FUNCTION_BLOCK Subestacao (* Subestacao / QGBT e geradores - ETE Tijuco Preto *)
  (* Standard: 61499-2 *)
  (* Version 1.2, 11/11/2026, Hidryco, Hidryco, 1.2: disjuntores ligados do PCE LODO (900) lidos pelo M262_Substacao na remota 1 do Lodo (.135): ${PATH}dj900_* e ${PATH}stsFalhaRemotaLODO -> IThis DJ_900_* e FALHA_REMOTA_LODO (PCE com logica invertida). 1.0: QGBT 440 V da ETE Tijuco Preto (unifilar HID-PE-DE-ETE-ELE-002): QTAM 1 (G2) -> 1Q1 -> barra A, QTAM 2 (G1) -> 1Q2 -> barra B, 1Q0 acoplamento. Disjuntores pelos DIs da remota 1 (A3/A4/A5 TM3DI32K do PCE SUBESTACAO) publicados por IO_DI32 em ${PATH}dj<nome>, ${PATH}mp<sinal>_1q<n> e ${PATH}stsFalhaRemota1. Geradores pelos Gerador_Generico internos GMG_G1 (QTAM 2) e GMG_G2 (QTAM 1). Cargas liberadas no gerador escolhidas na IHM (persistentes, padrao liberado): saidas HAB_* e stsPlantaNoGerador para os CATs de processo. v1.1: comandos de abrir/fechar dos Masterpact pela IHM (fpComandos) com intertravamentos, publicados em ${PATH}cmdAbrir1q1 ... ${PATH}cmdFechar1q2 para o IO_DQ32 do A8 TM3DQ32TK da remota 1 (word 0 b05..b10, escrita pelo M262_Substacao); reservas no unifilar. *)
  PACKAGE Hidryco.HidrycoLib;
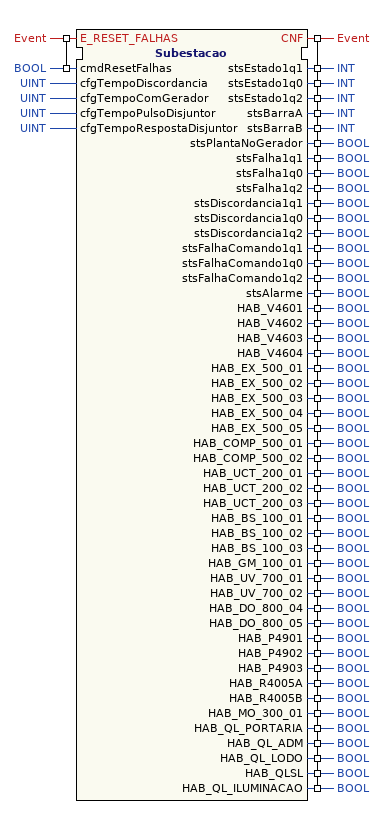
  EVENT_INPUT
    E_RESET_FALHAS WITH cmdResetFalhas; (* Reconhecimento pelo processo com cmdResetFalhas = TRUE *)
  END_EVENT
  EVENT_OUTPUT
    CNF WITH stsEstado1q1, stsEstado1q0, stsEstado1q2, stsBarraA, stsBarraB, stsPlantaNoGerador, stsFalha1q1, stsFalha1q0, stsFalha1q2, stsDiscordancia1q1, stsDiscordancia1q0, stsDiscordancia1q2, stsFalhaComando1q1, stsFalhaComando1q0, stsFalhaComando1q2, stsAlarme, HAB_V4601, HAB_V4602, HAB_V4603, HAB_V4604, HAB_EX_500_01, HAB_EX_500_02, HAB_EX_500_03, HAB_EX_500_04, HAB_EX_500_05, HAB_COMP_500_01, HAB_COMP_500_02, HAB_UCT_200_01, HAB_UCT_200_02, HAB_UCT_200_03, HAB_BS_100_01, HAB_BS_100_02, HAB_BS_100_03, HAB_GM_100_01, HAB_UV_700_01, HAB_UV_700_02, HAB_DO_800_04, HAB_DO_800_05, HAB_P4901, HAB_P4902, HAB_P4903, HAB_R4005A, HAB_R4005B, HAB_MO_300_01, HAB_QL_PORTARIA, HAB_QL_ADM, HAB_QL_LODO, HAB_QLSL, HAB_QL_ILUMINACAO; (* Estados do QGBT e cargas liberadas no gerador (so na mudanca) *)
  END_EVENT
  VAR_INPUT
    cmdResetFalhas : BOOL; (* TRUE = reconhecimento (com o evento E_RESET_FALHAS) *)
    cfgTempoDiscordancia : UINT := 5; (* Tempo (s) com aberto/fechado discordantes para o aviso de posicao indefinida *)
    cfgTempoComGerador : UINT := 10; (* Tempo (s) sem comunicacao com os AGC 150 para confirmar a falha *)
    cfgTempoPulsoDisjuntor : UINT := 1; (* Tempo (s) do pulso de abrir/fechar dos Masterpact (o pulso acaba antes se o disjuntor mudar de estado) *)
    cfgTempoRespostaDisjuntor : UINT := 5; (* Tempo (s) para o Masterpact mudar de estado depois do comando (senao: aviso de sem resposta) *)
  END_VAR
  VAR_OUTPUT
    stsEstado1q1 : INT; (* Disjuntor 1Q1: 0 indefinido (sem comunicacao), 1 aberto, 2 fechado, 3 discordante *)
    stsEstado1q0 : INT; (* Disjuntor 1Q0: 0 indefinido (sem comunicacao), 1 aberto, 2 fechado, 3 discordante *)
    stsEstado1q2 : INT; (* Disjuntor 1Q2: 0 indefinido (sem comunicacao), 1 aberto, 2 fechado, 3 discordante *)
    stsBarraA : INT; (* Fonte da barra A (1Q1): 0 sem alimentacao, 1 rede, 2 gerador, 3 indefinida *)
    stsBarraB : INT; (* Fonte da barra B (1Q2): 0 sem alimentacao, 1 rede, 2 gerador, 3 indefinida *)
    stsPlantaNoGerador : BOOL; (* Alguma QTAM com o disjuntor do gerador fechado (planta nos geradores) *)
    stsFalha1q1 : BOOL; (* Disjuntor 1Q1 em falha (desarmado) *)
    stsFalha1q0 : BOOL; (* Disjuntor 1Q0 em falha (desarmado) *)
    stsFalha1q2 : BOOL; (* Disjuntor 1Q2 em falha (desarmado) *)
    stsDiscordancia1q1 : BOOL; (* Disjuntor 1Q1: posição indefinida (aberto e fechado discordantes) *)
    stsDiscordancia1q0 : BOOL; (* Disjuntor 1Q0: posição indefinida (aberto e fechado discordantes) *)
    stsDiscordancia1q2 : BOOL; (* Disjuntor 1Q2: posição indefinida (aberto e fechado discordantes) *)
    stsFalhaComando1q1 : BOOL; (* Disjuntor 1Q1 não respondeu ao comando de abrir/fechar *)
    stsFalhaComando1q0 : BOOL; (* Disjuntor 1Q0 não respondeu ao comando de abrir/fechar *)
    stsFalhaComando1q2 : BOOL; (* Disjuntor 1Q2 não respondeu ao comando de abrir/fechar *)
    stsAlarme : BOOL; (* Algum alarme do QGBT *)
    HAB_V4601 : BOOL; (* V4601 - Soprador 01 liberado para operar com a planta nos geradores *)
    HAB_V4602 : BOOL; (* V4602 - Soprador 02 liberado para operar com a planta nos geradores *)
    HAB_V4603 : BOOL; (* V4603 - Soprador 03 liberado para operar com a planta nos geradores *)
    HAB_V4604 : BOOL; (* V4604 - Soprador 04 liberado para operar com a planta nos geradores *)
    HAB_EX_500_01 : BOOL; (* 500-EX-01 - Exaustor 01 liberado para operar com a planta nos geradores *)
    HAB_EX_500_02 : BOOL; (* 500-EX-02 - Exaustor 02 liberado para operar com a planta nos geradores *)
    HAB_EX_500_03 : BOOL; (* 500-EX-03 - Exaustor 03 liberado para operar com a planta nos geradores *)
    HAB_EX_500_04 : BOOL; (* 500-EX-04 - Exaustor 04 liberado para operar com a planta nos geradores *)
    HAB_EX_500_05 : BOOL; (* 500-EX-05 - Exaustor 05 liberado para operar com a planta nos geradores *)
    HAB_COMP_500_01 : BOOL; (* 500-COMP-01 - Compressor 01 liberado para operar com a planta nos geradores *)
    HAB_COMP_500_02 : BOOL; (* 500-COMP-02 - Compressor 02 liberado para operar com a planta nos geradores *)
    HAB_UCT_200_01 : BOOL; (* 200-UCT-01 - Unid. compacta 01 liberado para operar com a planta nos geradores *)
    HAB_UCT_200_02 : BOOL; (* 200-UCT-02 - Unid. compacta 02 liberado para operar com a planta nos geradores *)
    HAB_UCT_200_03 : BOOL; (* 200-UCT-03 - Unid. compacta 03 liberado para operar com a planta nos geradores *)
    HAB_BS_100_01 : BOOL; (* 100-BS-01 - Bomba 01 liberado para operar com a planta nos geradores *)
    HAB_BS_100_02 : BOOL; (* 100-BS-02 - Bomba 02 liberado para operar com a planta nos geradores *)
    HAB_BS_100_03 : BOOL; (* 100-BS-03 - Bomba 03 liberado para operar com a planta nos geradores *)
    HAB_GM_100_01 : BOOL; (* 100-GM-01 - Grade mecanizada liberado para operar com a planta nos geradores *)
    HAB_UV_700_01 : BOOL; (* 700-UV-01 - Sistema UV 01 liberado para operar com a planta nos geradores *)
    HAB_UV_700_02 : BOOL; (* 700-UV-02 - Sistema UV 02 liberado para operar com a planta nos geradores *)
    HAB_DO_800_04 : BOOL; (* 800-DO-04 - Bomba dosadora 04 liberado para operar com a planta nos geradores *)
    HAB_DO_800_05 : BOOL; (* 800-DO-05 - Bomba dosadora 05 liberado para operar com a planta nos geradores *)
    HAB_P4901 : BOOL; (* P4901 - Bomba submersível 01 liberado para operar com a planta nos geradores *)
    HAB_P4902 : BOOL; (* P4902 - Bomba submersível 02 liberado para operar com a planta nos geradores *)
    HAB_P4903 : BOOL; (* P4903 - Bomba submersível 03 liberado para operar com a planta nos geradores *)
    HAB_R4005A : BOOL; (* R4005A - Bomba horizontal A liberado para operar com a planta nos geradores *)
    HAB_R4005B : BOOL; (* R4005B - Bomba horizontal B liberado para operar com a planta nos geradores *)
    HAB_MO_300_01 : BOOL; (* 300-MO-01 - Misturador 01 liberado para operar com a planta nos geradores *)
    HAB_QL_PORTARIA : BOOL; (* QL Portaria liberado para operar com a planta nos geradores *)
    HAB_QL_ADM : BOOL; (* QL Administração liberado para operar com a planta nos geradores *)
    HAB_QL_LODO : BOOL; (* QL Lodo liberado para operar com a planta nos geradores *)
    HAB_QLSL : BOOL; (* QL Sala de quadros liberado para operar com a planta nos geradores *)
    HAB_QL_ILUMINACAO : BOOL; (* QL Iluminação externa liberado para operar com a planta nos geradores *)
  END_VAR
  FBS
    IThis : Subestacao_HMI(QI := TRUE);
    plcStart1 : plcStart(Prio := 10);
    Logica : basicSubestacao;
    Tick : E_CYCLE(DT := T#1s);
    GMG_G2 : Gerador_Generico;
    GMG_G1 : Gerador_Generico;
    Campo01 : SYMLINKMULTIVARDST_65D63179E2618F5E(NAME1 := '$${PATH}djRES_A1', NAME2 := '$${PATH}djRES_A2', NAME3 := '$${PATH}djPCM_EEE_BRUTO', NAME4 := '$${PATH}djPCM_DESINFECCAO', NAME5 := '$${PATH}djQGBT_220V', QI := TRUE); {SET_ATTRIBUTE(Configuration.GenericFBType.InterfaceParams, Runtime.System#I:=5;VALUE${I$}:BOOL,BOOL,BOOL,BOOL,BOOL)}
    Campo02 : SYMLINKMULTIVARDST_65D63179E2618F5E(NAME1 := '$${PATH}djUCT_200_01', NAME2 := '$${PATH}djCOMP_500_02', NAME3 := '$${PATH}djV4603', NAME4 := '$${PATH}djV4604', NAME5 := '$${PATH}djBANCO_CAPACITORES', QI := TRUE); {SET_ATTRIBUTE(Configuration.GenericFBType.InterfaceParams, Runtime.System#I:=5;VALUE${I$}:BOOL,BOOL,BOOL,BOOL,BOOL)}
    Campo03 : SYMLINKMULTIVARDST_65D63179E2618F5E(NAME1 := '$${PATH}djPCE_SUBESTACAO', NAME2 := '$${PATH}djCOMP_500_01', NAME3 := '$${PATH}djUCT_200_02', NAME4 := '$${PATH}djUCT_200_03', NAME5 := '$${PATH}djPCM_NEREDA', QI := TRUE); {SET_ATTRIBUTE(Configuration.GenericFBType.InterfaceParams, Runtime.System#I:=5;VALUE${I$}:BOOL,BOOL,BOOL,BOOL,BOOL)}
    Campo04 : SYMLINKMULTIVARDST_65D63179E2618F5E(NAME1 := '$${PATH}djPCM_LODO', NAME2 := '$${PATH}djCAP2', NAME3 := '$${PATH}djPCM_AGUA_REUSO', NAME4 := '$${PATH}djMO_500_01', NAME5 := '$${PATH}djV4601', QI := TRUE); {SET_ATTRIBUTE(Configuration.GenericFBType.InterfaceParams, Runtime.System#I:=5;VALUE${I$}:BOOL,BOOL,BOOL,BOOL,BOOL)}
    Campo05 : SYMLINKMULTIVARDST_65D63179E2618F5E(NAME1 := '$${PATH}djV4602', NAME2 := '$${PATH}djRES_B1', NAME3 := '$${PATH}djRES_B2', NAME4 := '$${PATH}djRES_B3', NAME5 := '$${PATH}djQGBT_220V_ENTRADA', QI := TRUE); {SET_ATTRIBUTE(Configuration.GenericFBType.InterfaceParams, Runtime.System#I:=5;VALUE${I$}:BOOL,BOOL,BOOL,BOOL,BOOL)}
    Campo06 : SYMLINKMULTIVARDST_65D63179E2618F5E(NAME1 := '$${PATH}djQL_ADM', NAME2 := '$${PATH}djQL_PORTARIA', NAME3 := '$${PATH}djQLSL', NAME4 := '$${PATH}djQL_ILUMINACAO', NAME5 := '$${PATH}djPCE_SOPRADORES', QI := TRUE); {SET_ATTRIBUTE(Configuration.GenericFBType.InterfaceParams, Runtime.System#I:=5;VALUE${I$}:BOOL,BOOL,BOOL,BOOL,BOOL)}
    Campo07 : SYMLINKMULTIVARDST_65D63179E2618F5E(NAME1 := '$${PATH}djQL_LODO', NAME2 := '$${PATH}djRES_C1', NAME3 := '$${PATH}djRES_C2', NAME4 := '$${PATH}djRES_C3', NAME5 := '$${PATH}djRES_C4', QI := TRUE); {SET_ATTRIBUTE(Configuration.GenericFBType.InterfaceParams, Runtime.System#I:=5;VALUE${I$}:BOOL,BOOL,BOOL,BOOL,BOOL)}
    Campo08 : SYMLINKMULTIVARDST_65D63179E2618F5E(NAME1 := '$${PATH}djRES_C5', NAME2 := '$${PATH}djRES_C6', NAME3 := '$${PATH}mpL_1q1', NAME4 := '$${PATH}mpR_1q1', NAME5 := '$${PATH}mpP_1q1', QI := TRUE); {SET_ATTRIBUTE(Configuration.GenericFBType.InterfaceParams, Runtime.System#I:=5;VALUE${I$}:BOOL,BOOL,BOOL,BOOL,BOOL)}
    Campo09 : SYMLINKMULTIVARDST_65D63179E2618F5E(NAME1 := '$${PATH}mpC_1q1', NAME2 := '$${PATH}mpSF_1q1', NAME3 := '$${PATH}mpAB_1q1', NAME4 := '$${PATH}mpFE_1q1', NAME5 := '$${PATH}mpL_1q0', QI := TRUE); {SET_ATTRIBUTE(Configuration.GenericFBType.InterfaceParams, Runtime.System#I:=5;VALUE${I$}:BOOL,BOOL,BOOL,BOOL,BOOL)}
    Campo10 : SYMLINKMULTIVARDST_65D63179E2618F5E(NAME1 := '$${PATH}mpR_1q0', NAME2 := '$${PATH}mpP_1q0', NAME3 := '$${PATH}mpC_1q0', NAME4 := '$${PATH}mpSF_1q0', NAME5 := '$${PATH}mpAB_1q0', QI := TRUE); {SET_ATTRIBUTE(Configuration.GenericFBType.InterfaceParams, Runtime.System#I:=5;VALUE${I$}:BOOL,BOOL,BOOL,BOOL,BOOL)}
    Campo11 : SYMLINKMULTIVARDST_65D63179E2618F5E(NAME1 := '$${PATH}mpFE_1q0', NAME2 := '$${PATH}mpL_1q2', NAME3 := '$${PATH}mpR_1q2', NAME4 := '$${PATH}mpP_1q2', NAME5 := '$${PATH}mpC_1q2', QI := TRUE); {SET_ATTRIBUTE(Configuration.GenericFBType.InterfaceParams, Runtime.System#I:=5;VALUE${I$}:BOOL,BOOL,BOOL,BOOL,BOOL)}
    Campo12 : SYMLINKMULTIVARDST_1559B0FF8170C9BA0(NAME1 := '$${PATH}mpSF_1q2', QI := TRUE); {SET_ATTRIBUTE(Configuration.GenericFBType.InterfaceParams, Runtime.System#I:=1;VALUE${I$}:BOOL)}
    Campo13 : SYMLINKMULTIVARDST_1559B0FF8170C9BA0(NAME1 := '$${PATH}mpAB_1q2', QI := TRUE); {SET_ATTRIBUTE(Configuration.GenericFBType.InterfaceParams, Runtime.System#I:=1;VALUE${I$}:BOOL)}
    Campo14 : SYMLINKMULTIVARDST_1559B0FF8170C9BA0(NAME1 := '$${PATH}mpFE_1q2', QI := TRUE); {SET_ATTRIBUTE(Configuration.GenericFBType.InterfaceParams, Runtime.System#I:=1;VALUE${I$}:BOOL)}
    Campo15 : SYMLINKMULTIVARDST_1559B0FF8170C9BA0(NAME1 := '$${PATH}stsFalhaRemota1', QI := TRUE); {SET_ATTRIBUTE(Configuration.GenericFBType.InterfaceParams, Runtime.System#I:=1;VALUE${I$}:BOOL)}
    AlarmeF1q1 : ALARM_BIT(TYPE := 1, ACKTYPE_1 := 2, ACTIVE := TRUE); {SET_ATTRIBUTE(HMI.AlarmText, Disjuntor 1Q1 desarmado (falha))}
    AlarmeF1q0 : ALARM_BIT(TYPE := 1, ACKTYPE_1 := 2, ACTIVE := TRUE); {SET_ATTRIBUTE(HMI.AlarmText, Disjuntor 1Q0 desarmado (falha))}
    AlarmeF1q2 : ALARM_BIT(TYPE := 1, ACKTYPE_1 := 2, ACTIVE := TRUE); {SET_ATTRIBUTE(HMI.AlarmText, Disjuntor 1Q2 desarmado (falha))}
    AlarmeD1q1 : ALARM_BIT(TYPE := 1, ACKTYPE_1 := 2, ACTIVE := TRUE); {SET_ATTRIBUTE(HMI.AlarmText, Disjuntor 1Q1 com posição indefinida (aberto e fechado discordantes))} {SET_ATTRIBUTE(HMI.AlarmClass, Warning)}
    AlarmeD1q0 : ALARM_BIT(TYPE := 1, ACKTYPE_1 := 2, ACTIVE := TRUE); {SET_ATTRIBUTE(HMI.AlarmText, Disjuntor 1Q0 com posição indefinida (aberto e fechado discordantes))} {SET_ATTRIBUTE(HMI.AlarmClass, Warning)}
    AlarmeD1q2 : ALARM_BIT(TYPE := 1, ACKTYPE_1 := 2, ACTIVE := TRUE); {SET_ATTRIBUTE(HMI.AlarmText, Disjuntor 1Q2 com posição indefinida (aberto e fechado discordantes))} {SET_ATTRIBUTE(HMI.AlarmClass, Warning)}
    AlarmeC1q1 : ALARM_BIT(TYPE := 1, ACKTYPE_1 := 2, ACTIVE := TRUE); {SET_ATTRIBUTE(HMI.AlarmText, Disjuntor 1Q1 não respondeu ao comando de abrir/fechar)} {SET_ATTRIBUTE(HMI.AlarmClass, Warning)}
    AlarmeC1q0 : ALARM_BIT(TYPE := 1, ACKTYPE_1 := 2, ACTIVE := TRUE); {SET_ATTRIBUTE(HMI.AlarmText, Disjuntor 1Q0 não respondeu ao comando de abrir/fechar)} {SET_ATTRIBUTE(HMI.AlarmClass, Warning)}
    AlarmeC1q2 : ALARM_BIT(TYPE := 1, ACKTYPE_1 := 2, ACTIVE := TRUE); {SET_ATTRIBUTE(HMI.AlarmText, Disjuntor 1Q2 não respondeu ao comando de abrir/fechar)} {SET_ATTRIBUTE(HMI.AlarmClass, Warning)}
    Campo16 : SYMLINKMULTIVARDST_65D63179E2618F5E(NAME1 := '$${PATH}djNER_PCE', NAME2 := '$${PATH}djNER_PCM', NAME3 := '$${PATH}djMO_300_01', NAME4 := '$${PATH}djR4005A', NAME5 := '$${PATH}djR4005B', QI := TRUE); {SET_ATTRIBUTE(Configuration.GenericFBType.InterfaceParams, Runtime.System#I:=5;VALUE${I$}:BOOL,BOOL,BOOL,BOOL,BOOL)}
    Campo17 : SYMLINKMULTIVARDST_65D63179E2618F5E(NAME1 := '$${PATH}djP4901', NAME2 := '$${PATH}djP4902', NAME3 := '$${PATH}djP4903', NAME4 := '$${PATH}djEEEB_PCE', NAME5 := '$${PATH}djEEEB_PCM', QI := TRUE); {SET_ATTRIBUTE(Configuration.GenericFBType.InterfaceParams, Runtime.System#I:=5;VALUE${I$}:BOOL,BOOL,BOOL,BOOL,BOOL)}
    Campo18 : SYMLINKMULTIVARDST_65D63179E2618F5E(NAME1 := '$${PATH}djCO_100_01', NAME2 := '$${PATH}djCO_100_02', NAME3 := '$${PATH}djCO_100_03', NAME4 := '$${PATH}djCO_100_04', NAME5 := '$${PATH}djGM_100_01_02', QI := TRUE); {SET_ATTRIBUTE(Configuration.GenericFBType.InterfaceParams, Runtime.System#I:=5;VALUE${I$}:BOOL,BOOL,BOOL,BOOL,BOOL)}
    Campo19 : SYMLINKMULTIVARDST_65D63179E2618F5E(NAME1 := '$${PATH}djMO_100_01', NAME2 := '$${PATH}djDES_PCE_DESLIGADO', NAME3 := '$${PATH}djDES_PCM_DESLIGADO', NAME4 := '$${PATH}djUV_700_01', NAME5 := '$${PATH}djUV_700_02', QI := TRUE); {SET_ATTRIBUTE(Configuration.GenericFBType.InterfaceParams, Runtime.System#I:=5;VALUE${I$}:BOOL,BOOL,BOOL,BOOL,BOOL)}
    Campo20 : SYMLINKMULTIVARDST_65D63179E2618F5E(NAME1 := '$${PATH}djVC_700_01', NAME2 := '$${PATH}djMO_700_01', NAME3 := '$${PATH}stsFalhaRemotaNER', NAME4 := '$${PATH}stsFalhaRemotaEEEB', NAME5 := '$${PATH}stsFalhaRemotaDES', QI := TRUE); {SET_ATTRIBUTE(Configuration.GenericFBType.InterfaceParams, Runtime.System#I:=5;VALUE${I$}:BOOL,BOOL,BOOL,BOOL,BOOL)}
    Lodo01 : SYMLINKMULTIVARDST_65D63179E2618F5E(NAME1 := '$${PATH}dj900_PCE_DESL', NAME2 := '$${PATH}dj900_PCM', NAME3 := '$${PATH}dj900_SO_01', NAME4 := '$${PATH}dj900_SO_02', NAME5 := '$${PATH}dj900_AD_01', QI := TRUE); {SET_ATTRIBUTE(Configuration.GenericFBType.InterfaceParams, Runtime.System#I:=5;VALUE${I$}:BOOL,BOOL,BOOL,BOOL,BOOL)}
    Lodo02 : SYMLINKMULTIVARDST_65D63179E2618F5E(NAME1 := '$${PATH}dj900_AD_02', NAME2 := '$${PATH}dj900_AD_03', NAME3 := '$${PATH}dj900_PP_01', NAME4 := '$${PATH}dj900_MN_01', NAME5 := '$${PATH}dj900_MN_02', QI := TRUE); {SET_ATTRIBUTE(Configuration.GenericFBType.InterfaceParams, Runtime.System#I:=5;VALUE${I$}:BOOL,BOOL,BOOL,BOOL,BOOL)}
    Lodo03 : SYMLINKMULTIVARDST_65D63179E2618F5E(NAME1 := '$${PATH}dj900_MN_03', NAME2 := '$${PATH}dj900_MN_04', NAME3 := '$${PATH}dj900_MN_05', NAME4 := '$${PATH}dj900_BO_01', NAME5 := '$${PATH}dj900_BO_02', QI := TRUE); {SET_ATTRIBUTE(Configuration.GenericFBType.InterfaceParams, Runtime.System#I:=5;VALUE${I$}:BOOL,BOOL,BOOL,BOOL,BOOL)}
    Lodo04 : SYMLINKMULTIVARDST_65D63179E2618F5E(NAME1 := '$${PATH}dj900_BO_03', NAME2 := '$${PATH}dj900_BR_01', NAME3 := '$${PATH}dj900_BR_02', NAME4 := '$${PATH}dj900_VA_01', NAME5 := '$${PATH}dj900_VA_02', QI := TRUE); {SET_ATTRIBUTE(Configuration.GenericFBType.InterfaceParams, Runtime.System#I:=5;VALUE${I$}:BOOL,BOOL,BOOL,BOOL,BOOL)}
    Lodo05 : SYMLINKMULTIVARDST_65D63179E2618F5E(NAME1 := '$${PATH}dj900_VE_01', NAME2 := '$${PATH}dj900_VE_02', NAME3 := '$${PATH}dj900_VA_06', NAME4 := '$${PATH}dj900_VA_07', NAME5 := '$${PATH}dj900_VA_08', QI := TRUE); {SET_ATTRIBUTE(Configuration.GenericFBType.InterfaceParams, Runtime.System#I:=5;VALUE${I$}:BOOL,BOOL,BOOL,BOOL,BOOL)}
    Lodo06 : SYMLINKMULTIVARDST_65D63179E2618F5E(NAME1 := '$${PATH}dj900_VA_09', NAME2 := '$${PATH}dj900_VA_10', NAME3 := '$${PATH}dj900_VA_11', NAME4 := '$${PATH}dj900_VA_12', NAME5 := '$${PATH}dj900_VA_13', QI := TRUE); {SET_ATTRIBUTE(Configuration.GenericFBType.InterfaceParams, Runtime.System#I:=5;VALUE${I$}:BOOL,BOOL,BOOL,BOOL,BOOL)}
    Lodo07 : SYMLINKMULTIVARDST_1559B0FF8170C9BA0(NAME1 := '$${PATH}dj900_VB_03', QI := TRUE); {SET_ATTRIBUTE(Configuration.GenericFBType.InterfaceParams, Runtime.System#I:=1;VALUE${I$}:BOOL)}
    Lodo08 : SYMLINKMULTIVARDST_1559B0FF8170C9BA0(NAME1 := '$${PATH}dj900_VB_04', QI := TRUE); {SET_ATTRIBUTE(Configuration.GenericFBType.InterfaceParams, Runtime.System#I:=1;VALUE${I$}:BOOL)}
    Lodo09 : SYMLINKMULTIVARDST_1559B0FF8170C9BA0(NAME1 := '$${PATH}stsFalhaRemotaLODO', QI := TRUE); {SET_ATTRIBUTE(Configuration.GenericFBType.InterfaceParams, Runtime.System#I:=1;VALUE${I$}:BOOL)}
    ComandoMP1 : SYMLINKMULTIVARSRC_151ACB50A2F8223B2(NAME1 := '$${PATH}cmdAbrir1q1', NAME2 := '$${PATH}cmdFechar1q1', NAME3 := '$${PATH}cmdAbrir1q0', QI := TRUE); {SET_ATTRIBUTE(Configuration.GenericFBType.InterfaceParams, Runtime.System#I:=3;VALUE${I$}:BOOL,BOOL,BOOL)}
    ComandoMP2 : SYMLINKMULTIVARSRC_151ACB50A2F8223B2(NAME1 := '$${PATH}cmdFechar1q0', NAME2 := '$${PATH}cmdAbrir1q2', NAME3 := '$${PATH}cmdFechar1q2', QI := TRUE); {SET_ATTRIBUTE(Configuration.GenericFBType.InterfaceParams, Runtime.System#I:=3;VALUE${I$}:BOOL,BOOL,BOOL)}
  END_FBS
  EVENT_CONNECTIONS
    plcStart1.FIRST_INIT TO IThis.01386593433D80B1;
    plcStart1.REDO_INIT TO IThis.01386593433D80B1;
    IThis.A63ACB8A73158E88 TO Logica.F0DD93C6F39257DB;
    Logica.0C14AE8D21235D8D TO Tick.START;
    Logica.0C14AE8D21235D8D TO Campo01.INIT;
    Logica.0C14AE8D21235D8D TO Campo02.INIT;
    Logica.0C14AE8D21235D8D TO Campo03.INIT;
    Logica.0C14AE8D21235D8D TO Campo04.INIT;
    Logica.0C14AE8D21235D8D TO Campo05.INIT;
    Logica.0C14AE8D21235D8D TO Campo06.INIT;
    Logica.0C14AE8D21235D8D TO Campo07.INIT;
    Logica.0C14AE8D21235D8D TO Campo08.INIT;
    Logica.0C14AE8D21235D8D TO Campo09.INIT;
    Logica.0C14AE8D21235D8D TO Campo10.INIT;
    Logica.0C14AE8D21235D8D TO Campo11.INIT;
    Logica.0C14AE8D21235D8D TO Campo12.INIT;
    Logica.0C14AE8D21235D8D TO Campo13.INIT;
    Logica.0C14AE8D21235D8D TO Campo14.INIT;
    Logica.0C14AE8D21235D8D TO Campo15.INIT;
    Logica.0C14AE8D21235D8D TO AlarmeF1q1.INIT;
    AlarmeF1q1.INITO TO AlarmeF1q1.REQ_INITDATA;
    AlarmeF1q1.CNF_INITDATA TO AlarmeF1q1.ACTIVATE;
    AlarmeF1q1.INITO TO AlarmeF1q0.INIT;
    AlarmeF1q0.INITO TO AlarmeF1q0.REQ_INITDATA;
    AlarmeF1q0.CNF_INITDATA TO AlarmeF1q0.ACTIVATE;
    AlarmeF1q0.INITO TO AlarmeF1q2.INIT;
    AlarmeF1q2.INITO TO AlarmeF1q2.REQ_INITDATA;
    AlarmeF1q2.CNF_INITDATA TO AlarmeF1q2.ACTIVATE;
    AlarmeF1q2.INITO TO AlarmeD1q1.INIT;
    AlarmeD1q1.INITO TO AlarmeD1q1.REQ_INITDATA;
    AlarmeD1q1.CNF_INITDATA TO AlarmeD1q1.ACTIVATE;
    AlarmeD1q1.INITO TO AlarmeD1q0.INIT;
    AlarmeD1q0.INITO TO AlarmeD1q0.REQ_INITDATA;
    AlarmeD1q0.CNF_INITDATA TO AlarmeD1q0.ACTIVATE;
    AlarmeD1q0.INITO TO AlarmeD1q2.INIT;
    AlarmeD1q2.INITO TO AlarmeD1q2.REQ_INITDATA;
    AlarmeD1q2.CNF_INITDATA TO AlarmeD1q2.ACTIVATE;
    AlarmeD1q2.INITO TO AlarmeC1q1.INIT;
    AlarmeC1q1.INITO TO AlarmeC1q1.REQ_INITDATA;
    AlarmeC1q1.CNF_INITDATA TO AlarmeC1q1.ACTIVATE;
    AlarmeC1q1.INITO TO AlarmeC1q0.INIT;
    AlarmeC1q0.INITO TO AlarmeC1q0.REQ_INITDATA;
    AlarmeC1q0.CNF_INITDATA TO AlarmeC1q0.ACTIVATE;
    AlarmeC1q0.INITO TO AlarmeC1q2.INIT;
    AlarmeC1q2.INITO TO AlarmeC1q2.REQ_INITDATA;
    AlarmeC1q2.CNF_INITDATA TO AlarmeC1q2.ACTIVATE;
    AlarmeC1q2.INITO TO plcStart1.ACK_FIRST;
    AlarmeC1q2.INITO TO IThis.BDA1C22C72F0DC6E;
    IThis.B3920EABC7A156A9 TO Logica.F60FCE8FB10EFC73;
    IThis.A53DBDA0C5474D6A TO Logica.9929BFFD9402DDB6;
    E_RESET_FALHAS TO Logica.823E1B5CF4461E23;
    Tick.EO TO Logica.13B54C4D85B7EA2E;
    Logica.705789F0F7F5D2C5 TO CNF;
    Logica.44A92DBC4672EE3B TO IThis.9B4185F7D8FD7429;
    IThis.557E557ECF0A66B6 TO Logica.3E677812C22D4014;
    Logica.0C14AE8D21235D8D TO ComandoMP1.INIT;
    Logica.88100C4D3B9DD5C4 TO ComandoMP1.REQ;
    Logica.0C14AE8D21235D8D TO ComandoMP2.INIT;
    Logica.88100C4D3B9DD5C4 TO ComandoMP2.REQ;
    Campo01.CNF TO IThis.9B4185F7D8FD7429;
    Campo02.CNF TO IThis.9B4185F7D8FD7429;
    Campo03.CNF TO IThis.9B4185F7D8FD7429;
    Campo04.CNF TO IThis.9B4185F7D8FD7429;
    Campo05.CNF TO IThis.9B4185F7D8FD7429;
    Campo06.CNF TO IThis.9B4185F7D8FD7429;
    Campo07.CNF TO IThis.9B4185F7D8FD7429;
    Campo08.CNF TO Logica.6567CC8D4EE5A245;
    Campo08.CNF TO IThis.9B4185F7D8FD7429;
    Campo09.CNF TO Logica.6567CC8D4EE5A245;
    Campo10.CNF TO Logica.6567CC8D4EE5A245;
    Campo11.CNF TO Logica.6567CC8D4EE5A245;
    Campo12.CNF TO Logica.6567CC8D4EE5A245;
    Campo13.CNF TO Logica.6567CC8D4EE5A245;
    Campo14.CNF TO Logica.6567CC8D4EE5A245;
    Campo15.CNF TO Logica.6567CC8D4EE5A245;
    GMG_G2.B61E80D27D776DFC TO Logica.87B2D1214C12141D;
    GMG_G2.B61E80D27D776DFC TO IThis.9B4185F7D8FD7429;
    IThis.A53DBDA0C5474D6A TO GMG_G2.7928A75A5088ACBD;
    E_RESET_FALHAS TO GMG_G2.7928A75A5088ACBD;
    GMG_G1.B61E80D27D776DFC TO Logica.87B2D1214C12141D;
    GMG_G1.B61E80D27D776DFC TO IThis.9B4185F7D8FD7429;
    IThis.A53DBDA0C5474D6A TO GMG_G1.7928A75A5088ACBD;
    E_RESET_FALHAS TO GMG_G1.7928A75A5088ACBD;
    Logica.AD81F22916A4D699 TO AlarmeF1q1.REQ;
    Logica.AD81F22916A4D699 TO AlarmeF1q0.REQ;
    Logica.AD81F22916A4D699 TO AlarmeF1q2.REQ;
    Logica.AD81F22916A4D699 TO AlarmeD1q1.REQ;
    Logica.AD81F22916A4D699 TO AlarmeD1q0.REQ;
    Logica.AD81F22916A4D699 TO AlarmeD1q2.REQ;
    Logica.AD81F22916A4D699 TO AlarmeC1q1.REQ;
    Logica.AD81F22916A4D699 TO AlarmeC1q0.REQ;
    Logica.AD81F22916A4D699 TO AlarmeC1q2.REQ;
    AlarmeF1q1.IND_1 TO IThis.9B4185F7D8FD7429;
    AlarmeF1q0.IND_1 TO IThis.9B4185F7D8FD7429;
    AlarmeF1q2.IND_1 TO IThis.9B4185F7D8FD7429;
    AlarmeD1q1.IND_1 TO IThis.9B4185F7D8FD7429;
    AlarmeD1q0.IND_1 TO IThis.9B4185F7D8FD7429;
    AlarmeD1q2.IND_1 TO IThis.9B4185F7D8FD7429;
    AlarmeC1q1.IND_1 TO IThis.9B4185F7D8FD7429;
    AlarmeC1q0.IND_1 TO IThis.9B4185F7D8FD7429;
    AlarmeC1q2.IND_1 TO IThis.9B4185F7D8FD7429;
    IThis.A53DBDA0C5474D6A TO AlarmeF1q1.ACK_C1;
    IThis.A53DBDA0C5474D6A TO AlarmeF1q0.ACK_C1;
    IThis.A53DBDA0C5474D6A TO AlarmeF1q2.ACK_C1;
    IThis.A53DBDA0C5474D6A TO AlarmeD1q1.ACK_C1;
    IThis.A53DBDA0C5474D6A TO AlarmeD1q0.ACK_C1;
    IThis.A53DBDA0C5474D6A TO AlarmeD1q2.ACK_C1;
    IThis.A53DBDA0C5474D6A TO AlarmeC1q1.ACK_C1;
    IThis.A53DBDA0C5474D6A TO AlarmeC1q0.ACK_C1;
    IThis.A53DBDA0C5474D6A TO AlarmeC1q2.ACK_C1;
    E_RESET_FALHAS TO AlarmeF1q1.ACK_C1;
    E_RESET_FALHAS TO AlarmeF1q0.ACK_C1;
    E_RESET_FALHAS TO AlarmeF1q2.ACK_C1;
    E_RESET_FALHAS TO AlarmeD1q1.ACK_C1;
    E_RESET_FALHAS TO AlarmeD1q0.ACK_C1;
    E_RESET_FALHAS TO AlarmeD1q2.ACK_C1;
    E_RESET_FALHAS TO AlarmeC1q1.ACK_C1;
    E_RESET_FALHAS TO AlarmeC1q0.ACK_C1;
    E_RESET_FALHAS TO AlarmeC1q2.ACK_C1;
    Logica.0C14AE8D21235D8D TO Campo16.INIT;
    Campo16.CNF TO IThis.9B4185F7D8FD7429;
    Logica.0C14AE8D21235D8D TO Campo17.INIT;
    Campo17.CNF TO IThis.9B4185F7D8FD7429;
    Logica.0C14AE8D21235D8D TO Campo18.INIT;
    Campo18.CNF TO IThis.9B4185F7D8FD7429;
    Logica.0C14AE8D21235D8D TO Campo19.INIT;
    Campo19.CNF TO IThis.9B4185F7D8FD7429;
    Logica.0C14AE8D21235D8D TO Campo20.INIT;
    Campo20.CNF TO IThis.9B4185F7D8FD7429;
    IThis.AD906B43DB32B2F8 TO Logica.E00B6991B4233CE8;
    IThis.91786E9747A5AF1B TO Logica.72E7C45E3F16D43D;
    IThis.C0A04441D90A26C6 TO Logica.C67BDF9EE3533293;
    IThis.F8CF6E0EF48DB29B TO Logica.595E0499F319E304;
    IThis.D54B14D55C063013 TO Logica.37499387BE57FB9C;
    IThis.42CF28208CFC0370 TO Logica.86D713EC07C37891;
    Logica.0C14AE8D21235D8D TO Lodo01.INIT;
    Lodo01.CNF TO IThis.9B4185F7D8FD7429;
    Logica.0C14AE8D21235D8D TO Lodo02.INIT;
    Lodo02.CNF TO IThis.9B4185F7D8FD7429;
    Logica.0C14AE8D21235D8D TO Lodo03.INIT;
    Lodo03.CNF TO IThis.9B4185F7D8FD7429;
    Logica.0C14AE8D21235D8D TO Lodo04.INIT;
    Lodo04.CNF TO IThis.9B4185F7D8FD7429;
    Logica.0C14AE8D21235D8D TO Lodo05.INIT;
    Lodo05.CNF TO IThis.9B4185F7D8FD7429;
    Logica.0C14AE8D21235D8D TO Lodo06.INIT;
    Lodo06.CNF TO IThis.9B4185F7D8FD7429;
    Logica.0C14AE8D21235D8D TO Lodo07.INIT;
    Lodo07.CNF TO IThis.9B4185F7D8FD7429;
    Logica.0C14AE8D21235D8D TO Lodo08.INIT;
    Lodo08.CNF TO IThis.9B4185F7D8FD7429;
    Logica.0C14AE8D21235D8D TO Lodo09.INIT;
    Lodo09.CNF TO IThis.9B4185F7D8FD7429;
  END_CONNECTIONS
  DATA_CONNECTIONS
    cfgTempoDiscordancia TO Logica.8C990B5C2FD24909;
    cfgTempoPulsoDisjuntor TO Logica.DD4A145AB55E3E82;
    cfgTempoRespostaDisjuntor TO Logica.744A23F794DF9B50;
    cmdResetFalhas TO Logica.6E4E631E3CCE89E2;
    cfgTempoComGerador TO GMG_G2.A410B91E1EF5ABA2;
    IThis.A4B8FB8677ED809C TO GMG_G2.19848145BDBC225E;
    GMG_G2.6A17B02D91A0D025 TO Logica.F40B2BFF770A4117;
    cfgTempoComGerador TO GMG_G1.A410B91E1EF5ABA2;
    IThis.A4B8FB8677ED809C TO GMG_G1.19848145BDBC225E;
    GMG_G1.6A17B02D91A0D025 TO Logica.A8803C88E516152D;
    Campo08.VALUE3 TO Logica.065477C347E2602C;
    Campo08.VALUE4 TO Logica.6FBEC1E5ECCA3874;
    Campo08.VALUE5 TO Logica.BCC87B7DB0119E13;
    Campo09.VALUE1 TO Logica.B7B198056E47289C;
    Campo09.VALUE2 TO Logica.2EB726DF525D8325;
    Campo09.VALUE3 TO Logica.76DD4ACCCAD07F91;
    Campo09.VALUE4 TO Logica.394C937F36C375C6;
    Campo09.VALUE5 TO Logica.D9C0B7637252BFAC;
    Campo10.VALUE1 TO Logica.2E33F99162E042B6;
    Campo10.VALUE2 TO Logica.48E50450CB3D0C81;
    Campo10.VALUE3 TO Logica.E45EB8FECC1FA9E4;
    Campo10.VALUE4 TO Logica.BFF0D2B31DF4374E;
    Campo10.VALUE5 TO Logica.F786AF3778AE631A;
    Campo11.VALUE1 TO Logica.000586804E10873D;
    Campo11.VALUE2 TO Logica.A90A3ECB125ABEF7;
    Campo11.VALUE3 TO Logica.D2844D138157228A;
    Campo11.VALUE4 TO Logica.CE5C20734596576E;
    Campo11.VALUE5 TO Logica.4A7111FBD61F99CE;
    Campo12.VALUE1 TO Logica.FACFB279B6DEAA8C;
    Campo13.VALUE1 TO Logica.FA5C14CCBC853FC7;
    Campo14.VALUE1 TO Logica.4BC3BB1293F9FBDE;
    Campo15.VALUE1 TO Logica.697402504175C39B;
    IThis.A49DF9844C61D026 TO Logica.7790FB996E34A50F;
    IThis.7DF7DF0127350B25 TO Logica.7C675CAD7ECE9CAE;
    IThis.1E75C26F37C04175 TO Logica.AD073A75439BCD3F;
    IThis.B4A0444CAEA4D1A6 TO Logica.1C58C750ADAFFB8D;
    IThis.EAC4C1EF3396CF05 TO Logica.2CC523736C76E209;
    IThis.1B21BD0DC1DEE349 TO Logica.D715D8E0A9ABBB07;
    IThis.98F440C9F3FA95D7 TO Logica.97081A98AFADD01C;
    IThis.6602639E11629D6A TO Logica.49CCAFDB9A9EB074;
    IThis.E71D50DEDD6FFE55 TO Logica.43A948136DCE906A;
    IThis.FE63B64AB87C4B66 TO Logica.D0BD9F60D08BBD1D;
    IThis.5489142ABCAABAF6 TO Logica.E9568CE9D1E184CD;
    IThis.B26E04769CA4882E TO Logica.D3E10E3648B70A9E;
    IThis.821EB5D7E791C714 TO Logica.E51D2D199E7E6DA3;
    IThis.13F650B4B20CAD30 TO Logica.092D56E4E9128DFF;
    IThis.D07E1CD7F0FD8F3D TO Logica.1550F9FE372176DC;
    IThis.8349228A3296D31B TO Logica.1BE22F2CAA170CAD;
    IThis.12EFE7ADF69BBAF1 TO Logica.60A40025609D9388;
    IThis.BC51424B486EA9FA TO Logica.ECDB1188ECF7F31B;
    IThis.3E03720186F6B8B4 TO Logica.8B7C83A062BEFDA6;
    IThis.1F72F37170B09B86 TO Logica.F585F77016D95C2A;
    IThis.CFA47B2CEBAC9DF5 TO Logica.F6E163DD85E8C55F;
    IThis.089857034819D352 TO Logica.01394094758A2B31;
    IThis.9064F938C9AC2A59 TO Logica.A1437B206D2D1247;
    IThis.E57B98A4497D31C1 TO Logica.BA1F8F2E3C393568;
    IThis.BE8F2E23CA76257B TO Logica.18C8D15491BE39F7;
    IThis.CD0B26C6013107D7 TO Logica.3CC5756FB770D61B;
    IThis.83DFCAD17CE085E4 TO Logica.EAE74B5D50AC23F7;
    IThis.EE81E9328A352B3B TO Logica.A754684D1774F264;
    IThis.62D42AC6D2F94586 TO Logica.FA116E94240DC36F;
    IThis.EF16D6E83472D1A1 TO Logica.E104FB97A1A0B09A;
    IThis.D8A7C20F42700B24 TO Logica.C47932E2565CC26D;
    IThis.C924E7FEDE79A00F TO Logica.955ECF78D67C4DF9;
    IThis.7FCD1D62A345B491 TO Logica.51FD70CCE0623138;
    IThis.A4B8FB8677ED809C TO Logica.B4F8B924E31359A1;
    IThis.D328525B197B17CB TO Logica.2CF5A6450291BD2C;
    Logica.82618CCEE38819DF TO ComandoMP1.VALUE1;
    Logica.E84C2E26BEE0CBD8 TO ComandoMP1.VALUE2;
    Logica.C01D66DF9D8D2B37 TO ComandoMP1.VALUE3;
    Logica.832E0476D93E3AB3 TO ComandoMP2.VALUE1;
    Logica.9C7D356999E24140 TO ComandoMP2.VALUE2;
    Logica.79D1A92C98189F87 TO ComandoMP2.VALUE3;
    Logica.1E69EF563D08B70A TO AlarmeF1q1.INP;
    Logica.F7D4AB497808F3EB TO AlarmeF1q0.INP;
    Logica.B0F14915CF2C7809 TO AlarmeF1q2.INP;
    Logica.592EF5C3E8B2B9FD TO AlarmeD1q1.INP;
    Logica.38C923E8FBD45478 TO AlarmeD1q0.INP;
    Logica.03139EE3DCF8782D TO AlarmeD1q2.INP;
    Logica.A61B09D63F370EB4 TO AlarmeC1q1.INP;
    Logica.F22ECF93013CE9A0 TO AlarmeC1q0.INP;
    Logica.BE9CBAB94EB8A2EC TO AlarmeC1q2.INP;
    Logica.CB2717BB76C89F56 TO stsEstado1q1;
    Logica.DA9419D5C7AA5DB3 TO stsEstado1q0;
    Logica.DFDB258CA97CCF9E TO stsEstado1q2;
    Logica.67FCF0CF94CE6434 TO stsBarraA;
    Logica.7900960E955E9B45 TO stsBarraB;
    Logica.F4BF7873F89E2578 TO stsPlantaNoGerador;
    Logica.3199FA5F3B5113A5 TO stsFalha1q1;
    Logica.9E350B5B0B15250A TO stsFalha1q0;
    Logica.2FA6B4B69E97CB81 TO stsFalha1q2;
    Logica.CDA8C144F8804259 TO stsDiscordancia1q1;
    Logica.9A580CA9D3A8ACA9 TO stsDiscordancia1q0;
    Logica.51AD3D0BCBA0D29F TO stsDiscordancia1q2;
    Logica.1CB488D6A7B45BD0 TO stsFalhaComando1q1;
    Logica.2FEAC3346B68E862 TO stsFalhaComando1q0;
    Logica.B720C4C18F3B0B83 TO stsFalhaComando1q2;
    Logica.7FF0CE8B8E26440C TO stsAlarme;
    Logica.21D2F882428D94F3 TO HAB_V4601;
    Logica.4BA2895B5E84852B TO HAB_V4602;
    Logica.0B6ADF853D305D47 TO HAB_V4603;
    Logica.BE34E4D2488C19E8 TO HAB_V4604;
    Logica.78A4F9EDC5C62C0C TO HAB_EX_500_01;
    Logica.1853F9A565699742 TO HAB_EX_500_02;
    Logica.E9F339DD43E61C92 TO HAB_EX_500_03;
    Logica.9C6435BC84B17E64 TO HAB_EX_500_04;
    Logica.BE7FE6C40B23C154 TO HAB_EX_500_05;
    Logica.CDE9A5680E80C4FC TO HAB_COMP_500_01;
    Logica.C423B287230633AC TO HAB_COMP_500_02;
    Logica.65AF809565D49EE4 TO HAB_UCT_200_01;
    Logica.FE43C0E5F49578C6 TO HAB_UCT_200_02;
    Logica.DFDF62B8B007BA30 TO HAB_UCT_200_03;
    Logica.A9DA853C672ACC03 TO HAB_BS_100_01;
    Logica.414CB46415187F9B TO HAB_BS_100_02;
    Logica.1A62A1CDE24C4BF5 TO HAB_BS_100_03;
    Logica.4F19BBB4DF5C103D TO HAB_GM_100_01;
    Logica.E6D53B29C9941104 TO HAB_UV_700_01;
    Logica.8013CE48BDBC119B TO HAB_UV_700_02;
    Logica.3D6D0C3D98EC3626 TO HAB_DO_800_04;
    Logica.73E4E38EB7FD8D14 TO HAB_DO_800_05;
    Logica.8C73844B4B959573 TO HAB_P4901;
    Logica.065415A90B86DB96 TO HAB_P4902;
    Logica.ECEAF09457E6C638 TO HAB_P4903;
    Logica.9A4F2AE3ADD5A02F TO HAB_R4005A;
    Logica.E96013B6D73D480C TO HAB_R4005B;
    Logica.FF26FAE248085DD1 TO HAB_MO_300_01;
    Logica.0BCE24EDE44554FA TO HAB_QL_PORTARIA;
    Logica.6EF58CFCE8899405 TO HAB_QL_ADM;
    Logica.1B43739444EC80C4 TO HAB_QL_LODO;
    Logica.1DCD400C037DE049 TO HAB_QLSL;
    Logica.9A4D494F76B758FC TO HAB_QL_ILUMINACAO;
    Campo01.VALUE1 TO IThis.596EE29105A45FA6;
    Campo01.VALUE2 TO IThis.45F9E7824916BC98;
    Campo01.VALUE3 TO IThis.AA8645BFAFB32BC9;
    Campo01.VALUE4 TO IThis.48A7FE9FF47A860D;
    Campo01.VALUE5 TO IThis.CCD7E78234D02ECE;
    Campo02.VALUE1 TO IThis.1270CD0D46E5DBE1;
    Campo02.VALUE2 TO IThis.87F9D8481AED82D4;
    Campo02.VALUE3 TO IThis.E661F967FD9F5842;
    Campo02.VALUE4 TO IThis.E95C9CCED4669773;
    Campo02.VALUE5 TO IThis.1CCEE621D5A72E0D;
    Campo03.VALUE1 TO IThis.525811933A8B0108;
    Campo03.VALUE2 TO IThis.BBB6F3F66F4A2157;
    Campo03.VALUE3 TO IThis.CE0A0EA52F933C29;
    Campo03.VALUE4 TO IThis.C4C9547C103F2643;
    Campo03.VALUE5 TO IThis.90AC1B67C96F5052;
    Campo04.VALUE1 TO IThis.6B4218E1FEB3CC79;
    Campo04.VALUE2 TO IThis.3712DDC6D8D3EF4A;
    Campo04.VALUE3 TO IThis.227AC21D2E93E1BF;
    Campo04.VALUE4 TO IThis.7648652FA873029B;
    Campo04.VALUE5 TO IThis.46F878B36A7B6DDD;
    Campo05.VALUE1 TO IThis.294F1C2FAA10CD3F;
    Campo05.VALUE2 TO IThis.605D8262C97CF729;
    Campo05.VALUE3 TO IThis.07FD230DFB59537F;
    Campo05.VALUE4 TO IThis.9BE0791E4227DC62;
    Campo05.VALUE5 TO IThis.4212351F67C78FF3;
    Campo06.VALUE1 TO IThis.8A6AD3A7FABAE5D1;
    Campo06.VALUE2 TO IThis.F762EDCBB2A78F45;
    Campo06.VALUE3 TO IThis.B82904E10ADB1EA3;
    Campo06.VALUE4 TO IThis.63C083BE8CD021FB;
    Campo06.VALUE5 TO IThis.4A7F4FF41597DC29;
    Campo07.VALUE1 TO IThis.B32E6D74DDA7B43A;
    Campo07.VALUE2 TO IThis.F9070970AC8E493A;
    Campo07.VALUE3 TO IThis.5E57006C5243DEBC;
    Campo07.VALUE4 TO IThis.1E37B3701F2AE226;
    Campo07.VALUE5 TO IThis.C1A7727AC4391022;
    Campo08.VALUE1 TO IThis.1DECAF3B8041CF27;
    Campo08.VALUE2 TO IThis.06C14CFF104482BE;
    Campo08.VALUE3 TO IThis.53C3DABD9672DE3F;
    Campo08.VALUE4 TO IThis.689BB1D3AC7A41D3;
    Campo08.VALUE5 TO IThis.D20049285A015725;
    Campo09.VALUE1 TO IThis.E81BE34AA05C5FBC;
    Campo09.VALUE2 TO IThis.350A4556E033D996;
    Campo09.VALUE5 TO IThis.9324D3A35375BADD;
    Campo10.VALUE1 TO IThis.873917FCA39E9FBE;
    Campo10.VALUE2 TO IThis.A612D03EDB3893BA;
    Campo10.VALUE3 TO IThis.D7E90ABA46BFA30E;
    Campo10.VALUE4 TO IThis.65DE5BE29C3C6131;
    Campo11.VALUE2 TO IThis.516E2910DFDD3665;
    Campo11.VALUE3 TO IThis.C375B7500AF8F5AD;
    Campo11.VALUE4 TO IThis.E3D17EF6F94BC74A;
    Campo11.VALUE5 TO IThis.D75B9FE6DE273C97;
    Campo12.VALUE1 TO IThis.D9C2FCCE62482B9A;
    Logica.CB2717BB76C89F56 TO IThis.BFEF898BE0511AE2;
    Logica.DA9419D5C7AA5DB3 TO IThis.98228BCDCC840B54;
    Logica.DFDB258CA97CCF9E TO IThis.5D56376579824383;
    Logica.67FCF0CF94CE6434 TO IThis.9E616DFC8D419447;
    Logica.7900960E955E9B45 TO IThis.8ACA15A20BDBF7EB;
    Logica.F4BF7873F89E2578 TO IThis.1B54C923B1CDB894;
    Campo15.VALUE1 TO IThis.24539C3AA2E83C47;
    GMG_G2.E607B5D65C774239 TO IThis.2E232C8392047708;
    GMG_G1.E607B5D65C774239 TO IThis.8090C8ED7C739DA3;
    GMG_G2.36AA02DF41051BAE TO IThis.1C891AA8DE6C4BFA;
    GMG_G1.36AA02DF41051BAE TO IThis.A04D304DCB1237A3;
    Logica.3199FA5F3B5113A5 TO IThis.0918E781740BFEEA;
    Logica.9E350B5B0B15250A TO IThis.F92674128CE8CE3C;
    Logica.2FA6B4B69E97CB81 TO IThis.9EE286C30D8DFD30;
    Logica.CDA8C144F8804259 TO IThis.93D475BF12719D66;
    Logica.9A580CA9D3A8ACA9 TO IThis.91DDDA71FE07A4E4;
    Logica.51AD3D0BCBA0D29F TO IThis.AAF0FAFDC7318CE0;
    Logica.1CB488D6A7B45BD0 TO IThis.79DD30B6EE021385;
    Logica.2FEAC3346B68E862 TO IThis.CB13A4C3ECAB260E;
    Logica.B720C4C18F3B0B83 TO IThis.6BE9EFC349A5D717;
    Logica.7FF0CE8B8E26440C TO IThis.85BED64DAA5E11C2;
    AlarmeF1q1.STATE_1 TO IThis.FBB32CFEEB2984DB;
    AlarmeF1q0.STATE_1 TO IThis.A71980BA56FC1CA0;
    AlarmeF1q2.STATE_1 TO IThis.B7EDF92D9560FDCA;
    AlarmeD1q1.STATE_1 TO IThis.0E1115BC4586C784;
    AlarmeD1q0.STATE_1 TO IThis.81AA7E50837D0AA4;
    AlarmeD1q2.STATE_1 TO IThis.40D86301893F3808;
    AlarmeC1q1.STATE_1 TO IThis.D6C986E35428EBC6;
    AlarmeC1q0.STATE_1 TO IThis.8C5C0CFF9E687FB2;
    AlarmeC1q2.STATE_1 TO IThis.6F85A52703A90075;
    Logica.D4E6388462E7070F TO IThis.51F3EECFC2110999;
    Logica.A0E35D1BB888A41D TO IThis.D0890CAF84480CCB;
    Logica.5A13984C5426C09A TO IThis.A2E371E74A6D47DF;
    Logica.CEFD3DC03D34D588 TO IThis.2D34900FFEBD9D67;
    Logica.4BAA35629E3CE6D0 TO IThis.CDB2B1C8D5C85226;
    Logica.8448BF8C1FCFD143 TO IThis.A6AE7EFA06A3684A;
    Logica.82618CCEE38819DF TO IThis.69483FE2E5DF433D;
    Logica.E84C2E26BEE0CBD8 TO IThis.58BE24B4AA8027FB;
    Logica.C01D66DF9D8D2B37 TO IThis.E5722FA7DF5CC4D5;
    Logica.832E0476D93E3AB3 TO IThis.18F792987566CE93;
    Logica.9C7D356999E24140 TO IThis.8E9F9CC231F1E34E;
    Logica.79D1A92C98189F87 TO IThis.F2764C516734F69E;
    Campo16.VALUE1 TO IThis.438C0D512EB97B9B;
    Campo16.VALUE2 TO IThis.D4FA5B3503D81F60;
    Campo16.VALUE3 TO IThis.857CCDF4E0CA6BFF;
    Campo16.VALUE4 TO IThis.63B76AD0D8107316;
    Campo16.VALUE5 TO IThis.76ECD75E7BCAC3BB;
    Campo17.VALUE1 TO IThis.45182DBF833B2661;
    Campo17.VALUE2 TO IThis.31F3A75D0C420C2C;
    Campo17.VALUE3 TO IThis.45112A3ED837A709;
    Campo17.VALUE4 TO IThis.BEC0D562D9236EDE;
    Campo17.VALUE5 TO IThis.62E398A490C6E7CA;
    Campo18.VALUE1 TO IThis.218C37A8CEC7D9CB;
    Campo18.VALUE2 TO IThis.B2EFD45DA7D8567A;
    Campo18.VALUE3 TO IThis.FD0AB6B6064A6BB0;
    Campo18.VALUE4 TO IThis.807C60DFDF9B1D34;
    Campo18.VALUE5 TO IThis.00606042F44B6636;
    Campo19.VALUE1 TO IThis.E37A0CFB51C1B827;
    Campo19.VALUE2 TO IThis.13A748A8D28A4926;
    Campo19.VALUE3 TO IThis.BAF1832AD07B033C;
    Campo19.VALUE4 TO IThis.26AA5FD004B208AF;
    Campo19.VALUE5 TO IThis.A2B95181FDFD5B87;
    Campo20.VALUE1 TO IThis.B054ECF246917636;
    Campo20.VALUE2 TO IThis.A2D107C92CF9E336;
    Campo20.VALUE3 TO IThis.ED60F77E117AFFE5;
    Campo20.VALUE4 TO IThis.2025666D77C7720C;
    Campo20.VALUE5 TO IThis.CFD6CDC749625C8A;
    Campo10.VALUE5 TO IThis.BE14C8E3A08C8666;
    Campo11.VALUE1 TO IThis.10C4CE673F7BDC3C;
    Campo09.VALUE3 TO IThis.E48B451401F5BBC5;
    Campo09.VALUE4 TO IThis.CBB765750A9DC70B;
    Campo13.VALUE1 TO IThis.848255A74DB7DC6D;
    Campo14.VALUE1 TO IThis.A3DDBCCC00EEF914;
    IThis.D2784D5AC7F3329D TO Logica.A367F1A895168A95;
    IThis.E58D37DBB6E4E2A0 TO Logica.242B879ED2446723;
    IThis.F384FB920A1B4FAD TO Logica.4621794953121717;
    IThis.D63D283E086C1625 TO Logica.621C7B35EA10B6F5;
    IThis.1463EB2C758A93FB TO Logica.5943FED7EE63C910;
    IThis.719A39E6AD840B6D TO Logica.F5DCE484B86495C1;
    Lodo01.VALUE1 TO IThis.B10C785E4683C1B6;
    Lodo01.VALUE2 TO IThis.1373ADB1D39EE182;
    Lodo01.VALUE3 TO IThis.448500E7DB550F95;
    Lodo01.VALUE4 TO IThis.8B8DD3B440CE42AC;
    Lodo01.VALUE5 TO IThis.D1C0BB941BF28EBB;
    Lodo02.VALUE1 TO IThis.4670EA26F25B5E3D;
    Lodo02.VALUE2 TO IThis.69A1461F54F625C6;
    Lodo02.VALUE3 TO IThis.7730CDE381FE264D;
    Lodo02.VALUE4 TO IThis.E02537D078F276D5;
    Lodo02.VALUE5 TO IThis.8E5083F6A4B4387A;
    Lodo03.VALUE1 TO IThis.0CF8CC05DB652F80;
    Lodo03.VALUE2 TO IThis.6DB9CC4795BCA41F;
    Lodo03.VALUE3 TO IThis.B8564152FA1B04B7;
    Lodo03.VALUE4 TO IThis.97824558375F0E5B;
    Lodo03.VALUE5 TO IThis.650D933F23BC0B22;
    Lodo04.VALUE1 TO IThis.30BEC7131C5A14A8;
    Lodo04.VALUE2 TO IThis.5DFC8535FB565FA4;
    Lodo04.VALUE3 TO IThis.ABA3CB28A43EDAD3;
    Lodo04.VALUE4 TO IThis.31A7371662CBE848;
    Lodo04.VALUE5 TO IThis.EE00E5FF917944D3;
    Lodo05.VALUE1 TO IThis.F22F25F79420BBEA;
    Lodo05.VALUE2 TO IThis.786C00DAB8635085;
    Lodo05.VALUE3 TO IThis.A47A1DDB4619794A;
    Lodo05.VALUE4 TO IThis.12363B0454BC23C4;
    Lodo05.VALUE5 TO IThis.74193D6A1F608DE7;
    Lodo06.VALUE1 TO IThis.F680C3FCE84DB3CD;
    Lodo06.VALUE2 TO IThis.B3C9BF39A7C6C290;
    Lodo06.VALUE3 TO IThis.38CEE3A723CF5518;
    Lodo06.VALUE4 TO IThis.397314465043FEA9;
    Lodo06.VALUE5 TO IThis.1181D2E87745533A;
    Lodo07.VALUE1 TO IThis.58E4ECC6FD4CD835;
    Lodo08.VALUE1 TO IThis.2884DE5F677AE328;
    Lodo09.VALUE1 TO IThis.536AA5CC2E6376A6;
  END_CONNECTIONS
END_FUNCTION_BLOCK
